{attribute 'qualified_only'}
{attribute 'to_string'}
TYPE E_ModeSelector :
(
    ModeNone := 0,
    FlipFlop := 1,
    Burst := 2,
    Open := 3,
    Close := 4,
    Home := 5
) UINT;
END_TYPE

(* stored: Version 1.1.0.1
   DUT E_ModeSelector: Id {f82f0162-029c-4006-a445-f48c61599328} *)
